FUNCTION_BLOCK FG_Transport

{region generated code}
VAR_INPUT
	Index01_B_Detect : FB_SensorBinary;
	Index01_B_Exit : FB_SensorBinary;
	Index01_Y_Lift : FB_Cylinder;
	Index01_Y_Stopper : FB_Cylinder;
	Index02_B_Detect : FB_SensorBinary;
	Index02_B_Exit : FB_SensorBinary;
	Index02_Y_Lift : FB_Cylinder;
	Index02_Y_Stopper : FB_Cylinder;
	Index03_B_Detect : FB_SensorBinary;
	Index03_B_Exit : FB_SensorBinary;
	Index03_Y_Lift : FB_Cylinder;
	Index03_Y_Stopper : FB_Cylinder;
	Index04_B_Detect : FB_SensorBinary;
	Index04_B_Exit : FB_SensorBinary;
	Index04_Y_Lift : FB_Cylinder;
	Index04_Y_Stopper : FB_Cylinder;
	Index05_B_Detect : FB_SensorBinary;
	Index05_B_Exit : FB_SensorBinary;
	Index05_Y_Lift : FB_Cylinder;
	Index05_Y_Stopper : FB_Cylinder;
	Lift01_B_Detect : FB_SensorBinary;
	Lift01_B_Exit : FB_SensorBinary;
	Lift01_M_Conveyor : FB_Drive;
	Lift01_Y_Lift : FB_Cylinder;
	Lift02_B_Detect : FB_SensorBinary;
	Lift02_B_Exit : FB_SensorBinary;
	Lift02_M_Conveyor : FB_Drive;
	Lift02_Y_Lift : FB_Cylinder;
	Stopper01_B_Detect : FB_SensorBinary;
	Stopper01_B_Exit : FB_SensorBinary;
	Stopper01_Y_Stopper : FB_Cylinder;
	Stopper02_B_Detect : FB_SensorBinary;
	Stopper02_B_Exit : FB_SensorBinary;
	Stopper02_Y_Stopper : FB_Cylinder;
	Stopper03_B_Detect : FB_SensorBinary;
	Stopper03_B_Exit : FB_SensorBinary;
	Stopper03_Y_Stopper : FB_Cylinder;
	Stopper04_B_Detect : FB_SensorBinary;
	Stopper04_B_Exit : FB_SensorBinary;
	Stopper04_Y_Stopper : FB_Cylinder;
	Transport01_M_Conveyor : FB_Drive;
	Transport02_M_Conveyor : FB_Drive;
END_VAR
{endregion}

{region generated code}
	InitRun();
	Index01_B_Detect();
	Index01_B_Exit();
	Index01_Y_Lift();
	Index01_Y_Stopper();
	Index02_B_Detect();
	Index02_B_Exit();
	Index02_Y_Lift();
	Index02_Y_Stopper();
	Index03_B_Detect();
	Index03_B_Exit();
	Index03_Y_Lift();
	Index03_Y_Stopper();
	Index04_B_Detect();
	Index04_B_Exit();
	Index04_Y_Lift();
	Index04_Y_Stopper();
	Index05_B_Detect();
	Index05_B_Exit();
	Index05_Y_Lift();
	Index05_Y_Stopper();
	Lift01_B_Detect();
	Lift01_B_Exit();
	Lift01_M_Conveyor();
	Lift01_Y_Lift();
	Lift02_B_Detect();
	Lift02_B_Exit();
	Lift02_M_Conveyor();
	Lift02_Y_Lift();
	Stopper01_B_Detect();
	Stopper01_B_Exit();
	Stopper01_Y_Stopper();
	Stopper02_B_Detect();
	Stopper02_B_Exit();
	Stopper02_Y_Stopper();
	Stopper03_B_Detect();
	Stopper03_B_Exit();
	Stopper03_Y_Stopper();
	Stopper04_B_Detect();
	Stopper04_B_Exit();
	Stopper04_Y_Stopper();
	Transport01_M_Conveyor();
	Transport02_M_Conveyor();
{endregion}

Mapping();

METHOD InitRun
{region generated code}
VAR_INST
	bInitRun : BOOL := TRUE;
END_VAR
{endregion}
{region generated code}
	IF NOT bInitRun THEN RETURN; END_IF
	bInitRun := FALSE;
{endregion}
END_METHOD

ACTION Mapping:
// ============================================================================
// FG_Transport twin <-> PLCSIM Advanced process image.
//
// Addresses: Siemens/_data/PLCTags_FG_Transport.xlsx.
//
// One byte per station, in the table's own order: Index01..05 on %I/%Q1003..1007,
// Stopper01..04 on 1008..1011, Lift01/02 on 1012/1013, Transport01/02 on
// 1014/1015. The bit positions repeat exactly per station type, so read one
// block and you have read them all.
//
// THE TWO GATES ARE NOT MAPPED HERE ANY MORE. FG_TS_Gate_1 / _2 keep their
// %I1001 / %I1002 addresses in this table, but the twin devices Y_Gate1 and
// Y_Gate2 live in FG_01 now - they are not members of this function block and
// assigning them here did not compile. They are mapped in FG_01's Mapping action,
// from these same addresses.
//
// Three things that are easy to get backwards:
//
//   * A STOPPER IS RETRACTED WHEN IT HOLDS THE PALLET. InHome %I1xxx.4 is
//     "Stopper geschlossen" and WorkPos %Q1xxx.2 is "Stopper oeffnen" - so
//     EXTENDING RELEASES. Nine authored Function entries in the twin say the
//     opposite and are known to be wrong; the table agrees with reality, not
//     with the twin's prose.
//   * A LIFT IS RETRACTED WHEN IT IS DOWN. InHome "Heber ist unten",
//     HomePos "Heber senken".
//   * ON A DRIVE, nControl.0 IS FORWARDS AND nControl.1 IS BACKWARDS. The table
//     names them: _Plus is "Antrieb vorwaerts", _Minus is "Antrieb rueckwaerts",
//     and Plus is always the LOWER address of the pair. THE PREVIOUS MAPPING HAD
//     ALL FOUR DRIVES INVERTED - it copied the Beckhoff side's channel order,
//     where the lower channel happens to be nControl.1, onto Siemens addresses
//     where the lower address is Plus. Every belt ran the wrong way.
// ============================================================================

// --- Index01 - detect, exit, lift and stopper on byte 1003 --------------
GVL_PLC.Inputs.I1003.0	:= Index01_B_Detect.bValue;
GVL_PLC.Inputs.I1003.1	:= Index01_B_Exit.bValue;
GVL_PLC.Inputs.I1003.2	:= Index01_Y_Lift.bRetracted;		// "Heber ist unten"
GVL_PLC.Inputs.I1003.3	:= Index01_Y_Lift.bExtended;		// "Heber ist oben"
GVL_PLC.Inputs.I1003.4	:= Index01_Y_Stopper.bRetracted;		// "Stopper geschlossen"
Index01_Y_Lift.bRetract	:= GVL_PLC.Outputs.Q1003.0;		// "Heber senken"
Index01_Y_Lift.bExtend	:= GVL_PLC.Outputs.Q1003.1;		// "Heber heben"
Index01_Y_Stopper.bExtend	:= GVL_PLC.Outputs.Q1003.2;		// "Stopper oeffnen"

// --- Index02 - detect, exit, lift and stopper on byte 1004 --------------
GVL_PLC.Inputs.I1004.0	:= Index02_B_Detect.bValue;
GVL_PLC.Inputs.I1004.1	:= Index02_B_Exit.bValue;
GVL_PLC.Inputs.I1004.2	:= Index02_Y_Lift.bRetracted;		// "Heber ist unten"
GVL_PLC.Inputs.I1004.3	:= Index02_Y_Lift.bExtended;		// "Heber ist oben"
GVL_PLC.Inputs.I1004.4	:= Index02_Y_Stopper.bRetracted;		// "Stopper geschlossen"
Index02_Y_Lift.bRetract	:= GVL_PLC.Outputs.Q1004.0;		// "Heber senken"
Index02_Y_Lift.bExtend	:= GVL_PLC.Outputs.Q1004.1;		// "Heber heben"
Index02_Y_Stopper.bExtend	:= GVL_PLC.Outputs.Q1004.2;		// "Stopper oeffnen"

// --- Index03 - detect, exit, lift and stopper on byte 1005 --------------
GVL_PLC.Inputs.I1005.0	:= Index03_B_Detect.bValue;
GVL_PLC.Inputs.I1005.1	:= Index03_B_Exit.bValue;
GVL_PLC.Inputs.I1005.2	:= Index03_Y_Lift.bRetracted;		// "Heber ist unten"
GVL_PLC.Inputs.I1005.3	:= Index03_Y_Lift.bExtended;		// "Heber ist oben"
GVL_PLC.Inputs.I1005.4	:= Index03_Y_Stopper.bRetracted;		// "Stopper geschlossen"
Index03_Y_Lift.bRetract	:= GVL_PLC.Outputs.Q1005.0;		// "Heber senken"
Index03_Y_Lift.bExtend	:= GVL_PLC.Outputs.Q1005.1;		// "Heber heben"
Index03_Y_Stopper.bExtend	:= GVL_PLC.Outputs.Q1005.2;		// "Stopper oeffnen"

// --- Index04 - detect, exit, lift and stopper on byte 1006 --------------
GVL_PLC.Inputs.I1006.0	:= Index04_B_Detect.bValue;
GVL_PLC.Inputs.I1006.1	:= Index04_B_Exit.bValue;
GVL_PLC.Inputs.I1006.2	:= Index04_Y_Lift.bRetracted;		// "Heber ist unten"
GVL_PLC.Inputs.I1006.3	:= Index04_Y_Lift.bExtended;		// "Heber ist oben"
GVL_PLC.Inputs.I1006.4	:= Index04_Y_Stopper.bRetracted;		// "Stopper geschlossen"
Index04_Y_Lift.bRetract	:= GVL_PLC.Outputs.Q1006.0;		// "Heber senken"
Index04_Y_Lift.bExtend	:= GVL_PLC.Outputs.Q1006.1;		// "Heber heben"
Index04_Y_Stopper.bExtend	:= GVL_PLC.Outputs.Q1006.2;		// "Stopper oeffnen"

// --- Index05 - detect, exit, lift and stopper on byte 1007 --------------
GVL_PLC.Inputs.I1007.0	:= Index05_B_Detect.bValue;
GVL_PLC.Inputs.I1007.1	:= Index05_B_Exit.bValue;
GVL_PLC.Inputs.I1007.2	:= Index05_Y_Lift.bRetracted;		// "Heber ist unten"
GVL_PLC.Inputs.I1007.3	:= Index05_Y_Lift.bExtended;		// "Heber ist oben"
GVL_PLC.Inputs.I1007.4	:= Index05_Y_Stopper.bRetracted;		// "Stopper geschlossen"
Index05_Y_Lift.bRetract	:= GVL_PLC.Outputs.Q1007.0;		// "Heber senken"
Index05_Y_Lift.bExtend	:= GVL_PLC.Outputs.Q1007.1;		// "Heber heben"
Index05_Y_Stopper.bExtend	:= GVL_PLC.Outputs.Q1007.2;		// "Stopper oeffnen"

// --- Stopper01 - detect, exit and stopper on byte 1008 --------------------
GVL_PLC.Inputs.I1008.0	:= Stopper01_B_Detect.bValue;
GVL_PLC.Inputs.I1008.1	:= Stopper01_B_Exit.bValue;
GVL_PLC.Inputs.I1008.4	:= Stopper01_Y_Stopper.bRetracted;		// "Stopper geschlossen"
Stopper01_Y_Stopper.bExtend	:= GVL_PLC.Outputs.Q1008.2;		// "Stopper oeffnen"

// --- Stopper02 - detect, exit and stopper on byte 1009 --------------------
GVL_PLC.Inputs.I1009.0	:= Stopper02_B_Detect.bValue;
GVL_PLC.Inputs.I1009.1	:= Stopper02_B_Exit.bValue;
GVL_PLC.Inputs.I1009.4	:= Stopper02_Y_Stopper.bRetracted;		// "Stopper geschlossen"
Stopper02_Y_Stopper.bExtend	:= GVL_PLC.Outputs.Q1009.2;		// "Stopper oeffnen"

// --- Stopper03 - detect, exit and stopper on byte 1010 --------------------
GVL_PLC.Inputs.I1010.0	:= Stopper03_B_Detect.bValue;
GVL_PLC.Inputs.I1010.1	:= Stopper03_B_Exit.bValue;
GVL_PLC.Inputs.I1010.4	:= Stopper03_Y_Stopper.bRetracted;		// "Stopper geschlossen"
Stopper03_Y_Stopper.bExtend	:= GVL_PLC.Outputs.Q1010.2;		// "Stopper oeffnen"

// --- Stopper04 - detect, exit and stopper on byte 1011 --------------------
GVL_PLC.Inputs.I1011.0	:= Stopper04_B_Detect.bValue;
GVL_PLC.Inputs.I1011.1	:= Stopper04_B_Exit.bValue;
GVL_PLC.Inputs.I1011.4	:= Stopper04_Y_Stopper.bRetracted;		// "Stopper geschlossen"
Stopper04_Y_Stopper.bExtend	:= GVL_PLC.Outputs.Q1011.2;		// "Stopper oeffnen"

// --- Lift01 - detect, exit, lift and carriage belt on byte 1012 --------
GVL_PLC.Inputs.I1012.0	:= Lift01_B_Detect.bValue;
GVL_PLC.Inputs.I1012.1	:= Lift01_B_Exit.bValue;
GVL_PLC.Inputs.I1012.2	:= Lift01_Y_Lift.bRetracted;		// "Heber ist unten"
GVL_PLC.Inputs.I1012.3	:= Lift01_Y_Lift.bExtended;		// "Heber ist oben"
Lift01_Y_Lift.bRetract	:= GVL_PLC.Outputs.Q1012.0;		// "Heber senken"
Lift01_Y_Lift.bExtend	:= GVL_PLC.Outputs.Q1012.1;		// "Heber heben"
Lift01_M_Conveyor.nControl.0	:= GVL_PLC.Outputs.Q1012.3;		// _Plus  "Antrieb vorwaerts"
Lift01_M_Conveyor.nControl.1	:= GVL_PLC.Outputs.Q1012.2;		// _Minus "Antrieb rueckwaerts"

// --- Lift02 - detect, exit, lift and carriage belt on byte 1013 --------
GVL_PLC.Inputs.I1013.0	:= Lift02_B_Detect.bValue;
GVL_PLC.Inputs.I1013.1	:= Lift02_B_Exit.bValue;
GVL_PLC.Inputs.I1013.2	:= Lift02_Y_Lift.bRetracted;		// "Heber ist unten"
GVL_PLC.Inputs.I1013.3	:= Lift02_Y_Lift.bExtended;		// "Heber ist oben"
Lift02_Y_Lift.bRetract	:= GVL_PLC.Outputs.Q1013.0;		// "Heber senken"
Lift02_Y_Lift.bExtend	:= GVL_PLC.Outputs.Q1013.1;		// "Heber heben"
Lift02_M_Conveyor.nControl.0	:= GVL_PLC.Outputs.Q1013.3;		// _Plus  "Antrieb vorwaerts"
Lift02_M_Conveyor.nControl.1	:= GVL_PLC.Outputs.Q1013.2;		// _Minus "Antrieb rueckwaerts"

// --- Transport01 - the level 1 circulation belt, byte 1014 -------------------
Transport01_M_Conveyor.nControl.0	:= GVL_PLC.Outputs.Q1014.1;		// _Plus  "Antrieb vorwaerts"
Transport01_M_Conveyor.nControl.1	:= GVL_PLC.Outputs.Q1014.0;		// _Minus "Antrieb rueckwaerts"

// --- Transport02 - the level 2 circulation belt, byte 1015 -------------------
Transport02_M_Conveyor.nControl.0	:= GVL_PLC.Outputs.Q1015.1;		// _Plus  "Antrieb vorwaerts"
Transport02_M_Conveyor.nControl.1	:= GVL_PLC.Outputs.Q1015.0;		// _Minus "Antrieb rueckwaerts"

// TODO: NO INPUT ADDRESS IN PLCTags_FG_Transport.xlsx for ANY of the four drives'
// running feedback. Every FB_Drive publishes nStatus.6 - "moving", written every
// scan - and none of the four has a tag for it, so the control PLC commands a belt
// and is never told whether it turned. A running belt is not a moving pallet, but
// a belt that never started is not either, and today the PLC cannot tell those
// apart. Add four input bits:
//   GVL_PLC.Inputs.I<n>.<b> := Lift01_M_Conveyor.nStatus.6;
//   GVL_PLC.Inputs.I<n>.<b> := Lift02_M_Conveyor.nStatus.6;
//   GVL_PLC.Inputs.I<n>.<b> := Transport01_M_Conveyor.nStatus.6;
//   GVL_PLC.Inputs.I<n>.<b> := Transport02_M_Conveyor.nStatus.6;
// nStatus.7 is NOT a health bit - it is a one second init pulse. Do not map it.

// TODO: NO Y_Stopper_InWork IN THE TABLE for any of the nine stoppers. Only the
// closed limit is published, so .bExtended goes nowhere and the PLC can see that
// a stopper has left the blocking position but never that it is fully clear. The
// Beckhoff side reads both limits on every stopper. Add %I1xxx.5 per station.
END_ACTION

END_FUNCTION_BLOCK

(* stored: Version 1.1.0.1, ProductVersion 3.1.4026.19
   POU FG_Transport: Id {1a228305-b0f2-406a-9e1d-b7bb3646ef17}, SpecialFunc None
   Method InitRun: Id {6e770fd6-c41f-4ee9-9c0d-3a96a1be5f92}
   Action Mapping: Id {62ee953e-c687-4d6b-a096-748c09bae4e3} *)
